Universal Robots URScript: T008_mistralai_Devstral-Small-2-24B-Instruct-2512_baseline_rep1_retry1.urscript

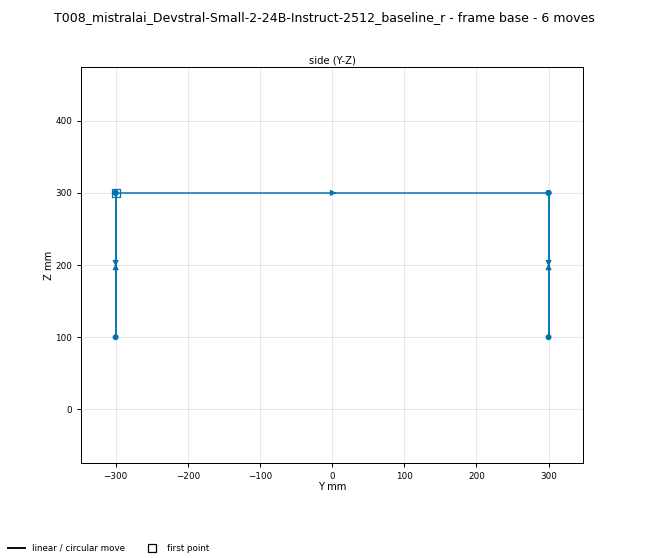
[picture p0: tool path of T008_mistralai_Devstral-Small-2-24B-Instruct-2512_baseline_rep1_retry1.urscript in frame base, 6 of 8 moves have a stored position in this frame; points joined in program order, loops and branches not executed]
def heavy_depalletizing():
    # Home position
    movej([0, -1.5708, 0, -1.5708, 0, 0], a=1.4, v=0.4, t=0, r=0)

    # Above pallet
    tool_zero_frame_acc = [1, 0, 0, 0, 0, 1, 0, 0, 0, 0, 0, 1, 0, 0, 0, 1]
    tool_zero_frame_vel = [1, 0, 0, 0, 0, 1, 0, 0, 0, 0, 0, 1, 0, 0, 0, 1]
    movel(p[0.5, -0.3, 0.3, 0, 3.14159, 0], a=1.4, v=0.4, t=0, r=0)

    # Descend to top layer
    movel(p[0.5, -0.3, 0.1, 0, 3.14159, 0], a=1.4, v=0.15, t=0, r=0)

    # Lift box
    movel(p[0.5, -0.3, 0.3, 0, 3.14159, 0], a=1.4, v=0.2, t=0, r=0)

    # Transit to conveyor
    movel(p[0.5, 0.3, 0.3, 0, 3.14159, 0], a=1.4, v=0.35, t=0, r=0)

    # Lower to conveyor
    movel(p[0.5, 0.3, 0.1, 0, 3.14159, 0], a=1.4, v=0.15, t=0, r=0)

    # Release box
    sleep(1.0)

    # Lift after release
    movel(p[0.5, 0.3, 0.3, 0, 3.14159, 0], a=1.4, v=0.2, t=0, r=0)

    # Return to home
    movej([0, -1.5708, 0, -1.5708, 0, 0], a=1.4, v=0.4, t=0, r=0)

heavy_depalletizing()
